TYPE ST_TriBlender :
STRUCT
	////Inputs
	bStartDisolving				: BOOL;
	
	sComponenetName			: STRING;
	sComponenetAmount		: STRING;
	tComponenetMixingTime	: TIME;
	tWaterCirculationTimeout: TIME;
	
	bLastComponent			: BOOL;	
	

	rMaxAllowedPressure		: REAL;
	rMinAllowedFlow			: REAL;
	bPumpOnFdbk				: BOOL;
	
	rPressure				: REAL;
	rFlow					: REAL;	
	rTemp					: REAL;
	
	
	///	outputs
	bError					: BOOL;
	sErrorDescription		: STRING;
	bDone					: BOOL;
	bComponenetMixDone		: BOOL;
	bDisolvingDone			: BOOL;
	

END_STRUCT
END_TYPE

(* stored: Version 1.1.0.1, ProductVersion 3.1.4024.13
   DUT ST_TriBlender: Id {402a54a6-73bc-4050-b13d-6e40fb7c3e37} *)
